(* IEC 61131-3 sources: kns-port-domestic/targets/astra/src/POUs/Model/FB_AnalogSensorSim, 2 files *)

(* ---- FB_AnalogSensorSim.decl.st ---- *)
// Назначение: датчик 4–20 мА в модели: ток = 4 + 16·(x − min)/(max − min) с насыщением
//             преобразователя на границах измерения NE 43 (3,8…20,5 мА), затем инъекция отказа
//             E_SimAiFault: обрыв (0 мА), токи отказа и выхода из диапазона SIM_MA_*, замерзание
//             (последний ток), принудительный ток. Неверная шкала или неконечное значение — ток
//             отказа снизу SIM_MA_FAIL_LOW (как у неисправного преобразователя).
// Автор:      kr0nsch
// Версия:     0.1.0
// Документ:   docs/DESIGN.md, раздел 11.2; docs/06_PMI.md, раздел 5.4
FUNCTION_BLOCK FB_AnalogSensorSim
VAR_INPUT
    rValue     : REAL;              // измеряемая величина, инж. ед.
    rRangeLo   : REAL;              // нижняя граница шкалы (4 мА)
    rRangeHi   : REAL;              // верхняя граница шкалы (20 мА)
    eFault     : E_SimAiFault;      // инъекция
    rForced_mA : REAL;              // ток при Forced
END_VAR
VAR_OUTPUT
    rCurrent_mA : REAL;             // ток в линии — вход модуля AI (GVL_IO.r<TAG>_mA)
END_VAR
VAR
    rMeas_mA : REAL;                // ток исправного преобразователя
END_VAR

(* ---- FB_AnalogSensorSim.impl.st ---- *)
// 1. Исправный преобразователь: линейная шкала и насыщение на границах измерения NE 43
IF PL.F_IsFinite(rIn := rValue) AND PL.F_IsFinite(rIn := rRangeLo) AND PL.F_IsFinite(rIn := rRangeHi)
   AND rRangeHi > rRangeLo THEN
    rMeas_mA := PL.GVL_Const.MA_ZERO + PL.GVL_Const.MA_SPAN * (rValue - rRangeLo) / (rRangeHi - rRangeLo);
    rMeas_mA := LIMIT(PL.GVL_Const.NE43_MEAS_LOW_MA, rMeas_mA, PL.GVL_Const.NE43_MEAS_HIGH_MA);
ELSE
    rMeas_mA := GVL_Const.SIM_MA_FAIL_LOW;
END_IF

// 2. Инъекция отказа (Freeze — ток прошлого вызова не меняется)
CASE eFault OF
    E_SimAiFault.WireBreak:
        rCurrent_mA := 0.0;
    E_SimAiFault.FailLow:
        rCurrent_mA := GVL_Const.SIM_MA_FAIL_LOW;
    E_SimAiFault.FailHigh:
        rCurrent_mA := GVL_Const.SIM_MA_FAIL_HIGH;
    E_SimAiFault.UnderRange:
        rCurrent_mA := GVL_Const.SIM_MA_UNDER_RANGE;
    E_SimAiFault.OverRange:
        rCurrent_mA := GVL_Const.SIM_MA_OVER_RANGE;
    E_SimAiFault.Freeze:
        // последнее значение тока
        ;
    E_SimAiFault.Forced:
        IF PL.F_IsFinite(rIn := rForced_mA) THEN
            rCurrent_mA := rForced_mA;
        ELSE
            rCurrent_mA := 0.0;
        END_IF
ELSE
    rCurrent_mA := rMeas_mA;
END_CASE
